// TIA Portal V20 export
// export: Created 2026-10-19T18:35:55.2771778Z, ExportSetting WithDefaults, DisplayName Totally Integrated Automation Portal, DisplayVersion V20 Update 6, DisplayName TIA Portal Openness, DisplayVersion V20 Update 6, DisplayName TIA Portal Version Control Interface, DisplayVersion V20 Update 6, DisplayName SINAMICS Startdrive Advanced, DisplayVersion V20 SP1, DisplayName SINAMICS Startdrive G130, G150, S120, S150, SINAMICS MV, G220, S200, S210, DisplayVersion V20 SP1, DisplayName SINAMICS Startdrive G110M, G120, G120C, G120D, G120P, G115D, DisplayVersion V20 SP1, DisplayName STEP 7 Professional, DisplayVersion V20 Update 6, DisplayName STEP 7 Safety, DisplayVersion V20 Update 2, DisplayName WinCC Basic/Comfort/Advanced, DisplayVersion V20 Update 6, DisplayName WinCC Unified, DisplayVersion V20 Update 6
DATA_BLOCK "Settings_DB"   // DB71
{ S7_Optimized_Access := 'TRUE' }
VERSION : 0.1
// stored: AutoNumber true, DBAccessibleFromOPCUA true, IsOnlyStoredInLoadMemory false, IsRetainMemResEnabled false, IsWriteProtectedInAS false, MemoryReserve 100
   VAR RETAIN
      VTD_Sys : Array[1..2] of "VTD_Settings";
      ECnv_Sys : Array[1..2] of "ECnv_Settings";
      LCnv_Sys : Array[1..2] of "Cnv_VTD_Settings";
      Shuttle_MQTT : "MQTT_Settings";
      System : "System_Settings";
   END_VAR
BEGIN
   VTD_Sys[1].ID := 1;
   VTD_Sys[2].ID := 2;
   VTD_Sys[1..2].Lowest_Level := 1;
   VTD_Sys[1..2].Highest_Level := 8;
   VTD_Sys[1..2].VTD_Max_Heigh := 16500;
   VTD_Sys[1].VTD_Min_Height := 55;
   VTD_Sys[2].VTD_Min_Height := 0;
   VTD_Sys[1..2].VTD_Level_Granularity := 20;
   VTD_Sys[1..2].Dft_Level_Offset_LE := 0;
   VTD_Sys[1..2].Dft_Level_Offset_AE := 0;
   VTD_Sys[1..2].Teach_Speed := 0;
   VTD_Sys[1..2].Creep_Speed := 3;
   VTD_Sys[1].Slow_Speed := 5;
   VTD_Sys[2].Slow_Speed := 15;
   VTD_Sys[1..2].Slow_Calib_Speed := 10;
   VTD_Sys[1..2].Loaded_Speed := 50;
   VTD_Sys[1..2].Shuttle_Speed := 50;
   VTD_Sys[1..2].Pallet_Speed := 100;
   VTD_Sys[1..2].Empty_Speed := 100;
   VTD_Sys[1..2].Dock_speed := 5;
   VTD_Sys[1..2].Manual_Speed := 15;
   VTD_Sys[1..2].Slowdown_Count_LE := 700;
   VTD_Sys[1].Creep_Count_LE := 60;
   VTD_Sys[2].Creep_Count_LE := 50;
   VTD_Sys[1..2].Slowdown_Count_AE := 700;
   VTD_Sys[1..2].Creep_Count_AE := 60;
   VTD_Sys[1..2].Encoder_Delta_W1 := 0.0;
   VTD_Sys[1..2].Encoder_Delta_W2 := 0.0;
   VTD_Sys[1..2].AE_Ratio := 0.0;
   VTD_Sys[1].Encoder_Delta_Warning := 80.0;
   VTD_Sys[2].Encoder_Delta_Warning := 50.0;
   VTD_Sys[1..2].Encoder_Delta_Error := 200.0;
   VTD_Sys[1..2].Transfer_Timeout_Up := 50;
   VTD_Sys[1..2].Transfer_Timeout_Down := 45;
   VTD_Sys[1..2].Lockpins_Timeout_Extend := 3000;
   VTD_Sys[1..2].Lockpins_Timeout_Retract := 3000;
   VTD_Sys[1].Level_Detect_Timeout := 500;
   VTD_Sys[2].Level_Detect_Timeout := 900;
   VTD_Sys[1..2].Teach_Timeout := 600;
   VTD_Sys[1].Chain_Slack_Timeout := 750;
   VTD_Sys[2].Chain_Slack_Timeout := 500;
   VTD_Sys[1].Level_Detect_LE := 3.0;
   VTD_Sys[2].Level_Detect_LE := 2.0;
   VTD_Sys[1..2].Acc_Range_1 := 60;
   VTD_Sys[1..2].Acc_Range_2 := 70;
   VTD_Sys[1..2].Acc_Range_3 := 80;
   VTD_Sys[1..2].Weight_Range_1 := 250;
   VTD_Sys[1..2].Weight_Range_2 := 500;
   VTD_Sys[1..2].Weight_Range_3 := 750;
   VTD_Sys[1].G120_Hardware_ID := 475;
   VTD_Sys[2].G120_Hardware_ID := 959;
   VTD_Sys[1].Teach_Values.Levels_LE[1] := 58.0;
   VTD_Sys[1].Teach_Values.Levels_LE[2] := 2525.0;
   VTD_Sys[1].Teach_Values.Levels_LE[3] := 4722.0;
   VTD_Sys[1].Teach_Values.Levels_LE[4] := 6927.0;
   VTD_Sys[1].Teach_Values.Levels_LE[5] := 9276.0;
   VTD_Sys[1].Teach_Values.Levels_LE[6] := 11627.0;
   VTD_Sys[1].Teach_Values.Levels_LE[7] := 13978.0;
   VTD_Sys[1].Teach_Values.Levels_LE[8] := 16325.0;
   VTD_Sys[2].Teach_Values.Levels_LE[1] := 63.0;
   VTD_Sys[2].Teach_Values.Levels_LE[2] := 2546.0;
   VTD_Sys[2].Teach_Values.Levels_LE[3] := 4744.0;
   VTD_Sys[2].Teach_Values.Levels_LE[4] := 6944.0;
   VTD_Sys[2].Teach_Values.Levels_LE[5] := 9291.0;
   VTD_Sys[2].Teach_Values.Levels_LE[6] := 11641.0;
   VTD_Sys[2].Teach_Values.Levels_LE[7] := 13993.0;
   VTD_Sys[2].Teach_Values.Levels_LE[8] := 16347.0;
   VTD_Sys[1].Teach_Values.Levels_AE[1..8] := 0;
   VTD_Sys[2].Teach_Values.Levels_AE[1..8] := 0;
   ECnv_Sys[1].ID := 120101;
   ECnv_Sys[2].ID := 120102;
   ECnv_Sys[1].Barcode_ID := 1;
   ECnv_Sys[2].Barcode_ID := 2;
   ECnv_Sys[1..2].Cnv_Level := 1;
   ECnv_Sys[1..2].TC_Time := 20;
   ECnv_Sys[1..2].Transfer_Time := 20;
   ECnv_Sys[1..2].Pallet_Align_Time := 20;
   ECnv_Sys[1..2].Slow_Speed := 10;
   ECnv_Sys[1..2].Full_Speed := 100;
   ECnv_Sys[1..2].Manual_Speed := 40;
   ECnv_Sys[1].G120_Hardware_ID := 488;
   ECnv_Sys[2].G120_Hardware_ID := 968;
   LCnv_Sys[1].Cnv_Level[2].Cnv1.ID := 100201;
   LCnv_Sys[1].Cnv_Level[3].Cnv1.ID := 100301;
   LCnv_Sys[1].Cnv_Level[4].Cnv1.ID := 100401;
   LCnv_Sys[1].Cnv_Level[5].Cnv1.ID := 100501;
   LCnv_Sys[1].Cnv_Level[6].Cnv1.ID := 100601;
   LCnv_Sys[2].Cnv_Level[2].Cnv1.ID := 100202;
   LCnv_Sys[2].Cnv_Level[3].Cnv1.ID := 100302;
   LCnv_Sys[2].Cnv_Level[4].Cnv1.ID := 100402;
   LCnv_Sys[2].Cnv_Level[5].Cnv1.ID := 100502;
   LCnv_Sys[2].Cnv_Level[6].Cnv1.ID := 100602;
   LCnv_Sys[1].Cnv_Level[2].Cnv1.Barcode_ID := 14;
   LCnv_Sys[1].Cnv_Level[3].Cnv1.Barcode_ID := 22;
   LCnv_Sys[1].Cnv_Level[4].Cnv1.Barcode_ID := 30;
   LCnv_Sys[1].Cnv_Level[5].Cnv1.Barcode_ID := 38;
   LCnv_Sys[1].Cnv_Level[6].Cnv1.Barcode_ID := 46;
   LCnv_Sys[2].Cnv_Level[2].Cnv1.Barcode_ID := 16;
   LCnv_Sys[2].Cnv_Level[3].Cnv1.Barcode_ID := 24;
   LCnv_Sys[2].Cnv_Level[4].Cnv1.Barcode_ID := 32;
   LCnv_Sys[2].Cnv_Level[5].Cnv1.Barcode_ID := 40;
   LCnv_Sys[2].Cnv_Level[6].Cnv1.Barcode_ID := 48;
   LCnv_Sys[1].Cnv_Level[2].Cnv1.Cnv_Level := 2;
   LCnv_Sys[1].Cnv_Level[3].Cnv1.Cnv_Level := 3;
   LCnv_Sys[1].Cnv_Level[4].Cnv1.Cnv_Level := 4;
   LCnv_Sys[1].Cnv_Level[5].Cnv1.Cnv_Level := 5;
   LCnv_Sys[1].Cnv_Level[6].Cnv1.Cnv_Level := 6;
   LCnv_Sys[2].Cnv_Level[2].Cnv1.Cnv_Level := 2;
   LCnv_Sys[2].Cnv_Level[3].Cnv1.Cnv_Level := 3;
   LCnv_Sys[2].Cnv_Level[4].Cnv1.Cnv_Level := 4;
   LCnv_Sys[2].Cnv_Level[5].Cnv1.Cnv_Level := 5;
   LCnv_Sys[2].Cnv_Level[6].Cnv1.Cnv_Level := 6;
   LCnv_Sys[1].Cnv_Level[2..6].Cnv1.TC_Time := 20;
   LCnv_Sys[2].Cnv_Level[2..6].Cnv1.TC_Time := 20;
   LCnv_Sys[1].Cnv_Level[2..6].Cnv1.Transfer_Time := 20;
   LCnv_Sys[2].Cnv_Level[2..6].Cnv1.Transfer_Time := 20;
   LCnv_Sys[1].Cnv_Level[2..6].Cnv1.Pallet_Align_Time := 20;
   LCnv_Sys[2].Cnv_Level[2..6].Cnv1.Pallet_Align_Time := 20;
   LCnv_Sys[1].Cnv_Level[2..6].Cnv1.Slow_Speed := 10;
   LCnv_Sys[2].Cnv_Level[2..6].Cnv1.Slow_Speed := 10;
   LCnv_Sys[1].Cnv_Level[2..6].Cnv1.Full_Speed := 86;
   LCnv_Sys[2].Cnv_Level[2..6].Cnv1.Full_Speed := 86;
   LCnv_Sys[1].Cnv_Level[2..6].Cnv1.Manual_Speed := 40;
   LCnv_Sys[2].Cnv_Level[2..6].Cnv1.Manual_Speed := 40;
   LCnv_Sys[1].Cnv_Level[2..6].Cnv1.Safety_stop_Timeout := 3000;
   LCnv_Sys[2].Cnv_Level[2..6].Cnv1.Safety_stop_Timeout := 3000;
   LCnv_Sys[1].Cnv_Level[2].Cnv1.G120_Hardware_ID := 551;
   LCnv_Sys[1].Cnv_Level[3].Cnv1.G120_Hardware_ID := 569;
   LCnv_Sys[1].Cnv_Level[4].Cnv1.G120_Hardware_ID := 581;
   LCnv_Sys[1].Cnv_Level[5].Cnv1.G120_Hardware_ID := 593;
   LCnv_Sys[1].Cnv_Level[6].Cnv1.G120_Hardware_ID := 605;
   LCnv_Sys[2].Cnv_Level[2].Cnv1.G120_Hardware_ID := 996;
   LCnv_Sys[2].Cnv_Level[3].Cnv1.G120_Hardware_ID := 1008;
   LCnv_Sys[2].Cnv_Level[4].Cnv1.G120_Hardware_ID := 1020;
   LCnv_Sys[2].Cnv_Level[5].Cnv1.G120_Hardware_ID := 1056;
   LCnv_Sys[2].Cnv_Level[6].Cnv1.G120_Hardware_ID := 1032;
   LCnv_Sys[1].Cnv_Level[2].Cnv2.ID := 110201;
   LCnv_Sys[1].Cnv_Level[3].Cnv2.ID := 110301;
   LCnv_Sys[1].Cnv_Level[4].Cnv2.ID := 110401;
   LCnv_Sys[1].Cnv_Level[5].Cnv2.ID := 110501;
   LCnv_Sys[1].Cnv_Level[6].Cnv2.ID := 110601;
   LCnv_Sys[2].Cnv_Level[2].Cnv2.ID := 110202;
   LCnv_Sys[2].Cnv_Level[3].Cnv2.ID := 110302;
   LCnv_Sys[2].Cnv_Level[4].Cnv2.ID := 110402;
   LCnv_Sys[2].Cnv_Level[5].Cnv2.ID := 110502;
   LCnv_Sys[2].Cnv_Level[6].Cnv2.ID := 110602;
   LCnv_Sys[1].Cnv_Level[2].Cnv2.Barcode_ID := 15;
   LCnv_Sys[1].Cnv_Level[3].Cnv2.Barcode_ID := 23;
   LCnv_Sys[1].Cnv_Level[4].Cnv2.Barcode_ID := 31;
   LCnv_Sys[1].Cnv_Level[5].Cnv2.Barcode_ID := 39;
   LCnv_Sys[1].Cnv_Level[6].Cnv2.Barcode_ID := 47;
   LCnv_Sys[2].Cnv_Level[2].Cnv2.Barcode_ID := 17;
   LCnv_Sys[2].Cnv_Level[3].Cnv2.Barcode_ID := 25;
   LCnv_Sys[2].Cnv_Level[4].Cnv2.Barcode_ID := 33;
   LCnv_Sys[2].Cnv_Level[5].Cnv2.Barcode_ID := 41;
   LCnv_Sys[2].Cnv_Level[6].Cnv2.Barcode_ID := 49;
   LCnv_Sys[1].Cnv_Level[2].Cnv2.Cnv_Level := 2;
   LCnv_Sys[1].Cnv_Level[3].Cnv2.Cnv_Level := 3;
   LCnv_Sys[1].Cnv_Level[4].Cnv2.Cnv_Level := 4;
   LCnv_Sys[1].Cnv_Level[5].Cnv2.Cnv_Level := 5;
   LCnv_Sys[1].Cnv_Level[6].Cnv2.Cnv_Level := 6;
   LCnv_Sys[2].Cnv_Level[2].Cnv2.Cnv_Level := 2;
   LCnv_Sys[2].Cnv_Level[3].Cnv2.Cnv_Level := 3;
   LCnv_Sys[2].Cnv_Level[4].Cnv2.Cnv_Level := 4;
   LCnv_Sys[2].Cnv_Level[5].Cnv2.Cnv_Level := 5;
   LCnv_Sys[2].Cnv_Level[6].Cnv2.Cnv_Level := 6;
   LCnv_Sys[1].Cnv_Level[2..6].Cnv2.TC_Time := 20;
   LCnv_Sys[2].Cnv_Level[2..6].Cnv2.TC_Time := 20;
   LCnv_Sys[1].Cnv_Level[2..6].Cnv2.Transfer_Time := 20;
   LCnv_Sys[2].Cnv_Level[2..6].Cnv2.Transfer_Time := 20;
   LCnv_Sys[1].Cnv_Level[2..6].Cnv2.Pallet_Align_Time := 20;
   LCnv_Sys[2].Cnv_Level[2..6].Cnv2.Pallet_Align_Time := 20;
   LCnv_Sys[1].Cnv_Level[2..6].Cnv2.Slow_Speed := 10;
   LCnv_Sys[2].Cnv_Level[2..6].Cnv2.Slow_Speed := 10;
   LCnv_Sys[1].Cnv_Level[2..6].Cnv2.Full_Speed := 86;
   LCnv_Sys[2].Cnv_Level[2..6].Cnv2.Full_Speed := 86;
   LCnv_Sys[1].Cnv_Level[2..6].Cnv2.Manual_Speed := 40;
   LCnv_Sys[2].Cnv_Level[2..6].Cnv2.Manual_Speed := 40;
   LCnv_Sys[1].Cnv_Level[2..6].Cnv2.Safety_stop_Timeout := 3000;
   LCnv_Sys[2].Cnv_Level[2..6].Cnv2.Safety_stop_Timeout := 3000;
   LCnv_Sys[1].Cnv_Level[2].Cnv2.G120_Hardware_ID := 641;
   LCnv_Sys[1].Cnv_Level[3].Cnv2.G120_Hardware_ID := 653;
   LCnv_Sys[1].Cnv_Level[4].Cnv2.G120_Hardware_ID := 665;
   LCnv_Sys[1].Cnv_Level[5].Cnv2.G120_Hardware_ID := 678;
   LCnv_Sys[1].Cnv_Level[6].Cnv2.G120_Hardware_ID := 690;
   LCnv_Sys[2].Cnv_Level[2].Cnv2.G120_Hardware_ID := 1092;
   LCnv_Sys[2].Cnv_Level[3].Cnv2.G120_Hardware_ID := 1104;
   LCnv_Sys[2].Cnv_Level[4].Cnv2.G120_Hardware_ID := 1116;
   LCnv_Sys[2].Cnv_Level[5].Cnv2.G120_Hardware_ID := 1128;
   LCnv_Sys[2].Cnv_Level[6].Cnv2.G120_Hardware_ID := 1140;
   Shuttle_MQTT.MQTT_Con_Params.hwId := 0;
   Shuttle_MQTT.MQTT_Con_Params.connId := 16#0001;
   Shuttle_MQTT.MQTT_Con_Params.broker := '10.44.116.9';
   Shuttle_MQTT.MQTT_Con_Params.port := 1883;
   Shuttle_MQTT.MQTT_Con_Params.tls.enableTls := FALSE;
   Shuttle_MQTT.MQTT_Con_Params.tls.validateServerIdentity := FALSE;
   Shuttle_MQTT.MQTT_Con_Params.tls.brokerCert := 0;
   Shuttle_MQTT.MQTT_Con_Params.tls.clientCert := 0;
   Shuttle_MQTT.MQTT_Con_Params.keepAlive := 60;
   Shuttle_MQTT.Client_ID := WSTRING#'PLC_1';
   Shuttle_MQTT.Username := WSTRING#'';
   Shuttle_MQTT.Password := WSTRING#'';
   Shuttle_MQTT.Timeout := 0;
   Shuttle_MQTT.QoS := 0;
   Shuttle_MQTT.Retain := TRUE;
   Shuttle_MQTT.Will_Topic := WSTRING#'';
   Shuttle_MQTT.Will_Msg_Length := 0;
   Shuttle_MQTT.Will_Msg_Payload[1..128] := 16#00;
   System.VTD_Count := 2;
   System.Level_Count := 6;
   System.Cnv_Count := 22;
   System.Shuttle_Count := 10;
   System.Shuttle_Interlock_Timeout := 999;
END_DATA_BLOCK
